Fanuc KAREL source: KA00200.KL

PROGRAM KA00200
%NOLOCKGROUP
VAR
  SRC: ARRAY[4] OF VECTOR
  DST: ARRAY[4] OF REAL
BEGIN
  DST = SRC
END KA00200
